Fanuc KAREL source: kb00071.KL

-- PROVISIONAL review KL for V1013-1; original PC SHA256 b98bbbef543c0bb84814f64262fe3f4adc1af79fb7e2db419d6d93f6a7af65a3
-- Incomplete behavior may be omitted. Consult companion uncertainty JSON. Do not deploy.
PROGRAM KB00071
%NOLOCKGROUP
VAR
  P1 : REAL
  RESULT : REAL
BEGIN
  -- UNRESOLVED_PC offsets 5-16; opcodes 2E,23
  -- UNRESOLVED_PC offsets 21-36; opcodes 27,22,76,23
  -- UNRESOLVED_PC offsets 41-45; opcodes 7F
END KB00071
